FUNCTION_BLOCK FB_ParameterHandler EXTENDS KOSTAL_AF2024_HMI_WinHMI.FB_Parameters_Base IMPLEMENTS I_Parameters_MainControl
VAR
END_VAR

PROPERTY airPressureMax : INT
GET
airPressureMax:= STRING_TO_INT(_getParameterValue(index:= E_Parameters.airPressureMax));
END_GET
END_PROPERTY

PROPERTY airPressureMin : INT
GET
airPressureMin:= STRING_TO_INT(_getParameterValue(index:= E_Parameters.airPressureMin));
END_GET
END_PROPERTY

{warning 'add property implementation'}
PROPERTY cylinderSensorTimeout : TIME
GET
cylinderSensorTimeout:= STRING_TO_TIME(_getParameterValue(index:= E_Parameters.cylinderTimeout));
END_GET
END_PROPERTY

METHOD FB_init : BOOL
VAR_INPUT
	bInitRetains 	: BOOL; // if TRUE, the retain variables are initialized (warm start / cold start)
	bInCopyCode 	: BOOL;  // if TRUE, the instance afterwards gets moved into the copy code (online change)
	ID_Name			: KOSTAL_AF2024_Core_Settings.T_MaxString;
	ID_Key			: DINT;
	CommonText		: KOSTAL_AF2024_Core_Text.I_Text;
	parameterPath	: KOSTAL_AF2024_Core_Settings.T_MaxString_UTF8;
	SystemTime		: KOSTAL_AF2024_Core_GetSystemTime.I_TimeSource;
END_VAR
_fullQualifiedFile:= parameterPath;
_I_getTime:= SystemTime;
END_METHOD

{warning 'add property implementation'}
PROPERTY isLoggerEnabled : BOOL
GET
isLoggerEnabled:= STRING_TO_BOOL(_getParameterValue(index:= E_Parameters.isLoggerEnabled));
END_GET
END_PROPERTY

{warning 'add property implementation'}
PROPERTY isNagaraEnable : BOOL
GET
isNagaraEnable:= STRING_TO_BOOL(_getParameterValue(index:= E_Parameters.isNagaraEnable));
END_GET
END_PROPERTY

{warning 'add property implementation'}
PROPERTY numberOfRetries : INT
GET
airPressureMax:= STRING_TO_INT(_getParameterValue(index:= E_Parameters.numberOfRetries));
END_GET
END_PROPERTY

END_FUNCTION_BLOCK

(* stored: Version 1.1.0.1, ProductVersion 3.1.4024.12
   POU FB_ParameterHandler: Id {de5c841e-3290-0e6b-0bfb-3f8135565583}, SpecialFunc None
   Folder I_Parameters_MainControl: Id {e90b4100-972e-05fd-04cc-db66b386c159}
   Folder Private: Id {c9d2c9b0-249c-055b-13da-628e2e99e886}
   Property airPressureMax: Id {d7cc16d0-eec9-0cac-341a-d31e5153d990}
   Get Get: Id {9af21b3c-cd52-023e-0123-7e5578ec07a4}
   Property airPressureMin: Id {5f3b26d9-3ff3-0b2f-1a8f-c3cbdea25a95}
   Get Get: Id {e7b034a8-1802-0e24-3e9b-d77c7099903a}
   Property cylinderSensorTimeout: Id {ea90df9f-98c5-475b-ab5f-3f8534cba318}
   Get Get: Id {4cb9fb38-069d-4044-b903-c8b5dc9d8e07}
   Method FB_init: Id {1651d52f-d2b9-09a9-2e7b-a3f01a6ad6da}
   Property isLoggerEnabled: Id {acdfb1c0-6703-466f-be43-1271096a24fb}
   Get Get: Id {5c7f0837-99b7-421c-b043-82c6bf719d4c}
   Property isNagaraEnable: Id {67c2fa63-96c7-4e1b-a61f-a2dbd242dfe2}
   Get Get: Id {f54bbad3-a054-41d9-b4cb-a58b61233e70}
   Property numberOfRetries: Id {38a0335f-7704-41b4-acc3-df5268f0ff89}
   Get Get: Id {3686a156-9dbf-4b17-8288-d74d68ac16b3} *)
